(* IEC 61131-3 sources: iolistgen/pytests/golden/gen_fixture/src/POUs/Generated/PRG_Devices, 2 files *)

(* ---- PRG_Devices.decl.st ---- *)
// AUTO-GENERATED by iolistgen 0.2.0 — не редактировать; источник: gen_fixture.csv
// SHA-256 перечня 3ace79e7a28b; генератор st-codesys
// Назначение: вызовы устройств plc-process-lib по перечню сигналов: входы из GVL_IO, выходы в GVL_IO, команды GVL_Hmi,
// Cfg и Retain — GVL_Persist (контракт plc-process-lib, разделы 1 и 20). Входы автоматики (xAutoRun, xAutoOpen,
// wInterlock, wPermit…, rSpeedSpAuto_pct, rPosSpAuto_pct) пишет логика станции до вызова PRG_Devices; ПИД-регуляторы
// (тип Pid) без сигналов ввода-вывода вызывает логика станции (контракт 17.3)
// Автор:      iolistgen (генератор по перечню сигналов); перечень gen_fixture.csv
// Версия:     iolistgen 0.2.0
// Документ:   docs/signal_list.md
PROGRAM PRG_Devices
VAR
END_VAR

(* ---- PRG_Devices.impl.st ---- *)
// AUTO-GENERATED by iolistgen 0.2.0 — не редактировать; источник: gen_fixture.csv
// SHA-256 перечня 3ace79e7a28b; генератор st-codesys
// Порядок: устройства, на которые ссылаются link_power и link_fb (PWR2, ZT201), вызываются раньше ссылающихся; дальше —
// по dev_no.
// Источник времени не привязан: устройства берут встроенное системное время (контракт 20).

// Команда HMI «Применить уставки проекта» (контракт 18.3, правило 2): Retain устройств не меняется
IF GVL_Hmi.xApplyProjectCfg THEN
    GVL_Hmi.xApplyProjectCfg := FALSE;
    PRG_ApplyProjectCfg();
END_IF

// --- dev_no 6: PWR2 — Напряжение на секции шин (DigitalInput) ---
GVL_Devices.fbPWR2(
    xIn           := GVL_IO.xPWR2,
    xChannelFault := FALSE,  // нет строки CHF
    stCmd         := GVL_Hmi.stPWR2Cmd,
    stCfg         := GVL_Persist.stPWR2Cfg);

// --- dev_no 32: ZT201 — Клапан рециркуляции: положение (AnalogInput) ---
GVL_Devices.fbZT201(
    rIn           := GVL_IO.rZT201_mA,
    xChannelFault := FALSE,  // нет строки CHF
    stCmd         := GVL_Hmi.stZT201Cmd,
    stCfg         := GVL_Persist.stZT201Cfg);

// --- dev_no 1: LT201 — Уровень в резервуаре чистой воды (AnalogInput) ---
GVL_Devices.fbLT201(
    rIn           := GVL_IO.rLT201_mA,
    xChannelFault := GVL_IO.xLT201_CHF,
    stCmd         := GVL_Hmi.stLT201Cmd,
    stCfg         := GVL_Persist.stLT201Cfg);

// --- dev_no 2: PT201 — Давление на всасе (AnalogInput) ---
GVL_Devices.fbPT201(
    rIn           := INT_TO_REAL(GVL_IO.iPT201),
    xChannelFault := NOT GVL_IO.xMbOk_RS485_1_S5,  // нет строки CHF: обмен со слейвом
    stCmd         := GVL_Hmi.stPT201Cmd,
    stCfg         := GVL_Persist.stPT201Cfg);

// --- dev_no 3: TE201 — Температура воды (AnalogInput) ---
GVL_Devices.fbTE201(
    rIn           := GVL_IO.rTE201,
    xChannelFault := FALSE,  // нет строки CHF
    stCmd         := GVL_Hmi.stTE201Cmd,
    stCfg         := GVL_Persist.stTE201Cfg);

// --- dev_no 4: LS201 — Поплавок «перелив» (DigitalInput) ---
GVL_Devices.fbLS201(
    xIn           := GVL_IO.xLS201,
    xChannelFault := GVL_IO.xLS201_CHF,
    stCmd         := GVL_Hmi.stLS201Cmd,
    stCfg         := GVL_Persist.stLS201Cfg);

// --- dev_no 5: ES201 — Кнопка аварийного останова на щите (DigitalInput) ---
GVL_Devices.fbES201(
    xIn           := GVL_IO.xES201,
    xChannelFault := NOT GVL_IO.xMbOk_RS485_1_S7,  // нет строки CHF: обмен со слейвом
    stCmd         := GVL_Hmi.stES201Cmd,
    stCfg         := GVL_Persist.stES201Cfg);

// --- dev_no 11: M201 — Насос промывки (Motor) ---
GVL_Devices.fbM201(
    xFbRun    := GVL_IO.xM201_FB,
    xExtFault := GVL_IO.xM201_FLT,
    xLocal    := GVL_IO.xM201_LOC,
    xPowerOk  := GVL_Devices.fbPWR2.xValue,  // link_power
    stCmd     := GVL_Hmi.stM201Cmd,
    stCfg     := GVL_Persist.stM201Cfg,
    stRetain  := GVL_Persist.stM201Retain);
GVL_IO.xM201_RUN := GVL_Devices.fbM201.xQRun;
GVL_IO.xM201_RST := GVL_Devices.fbM201.xQReset;

// --- dev_no 12: P201 — Насос Н1 (MotorVfd) ---
// ПЧ: xCommOk, xVfd*, rSpeedAct_pct и rSpeedRef_pct — через адаптер приложения (GVL_IO.xP201_…)
GVL_Devices.fbP201(
    xExtFault     := GVL_IO.xP201_FLT,
    xLocal        := GVL_IO.xP201_LOC,
    xPowerOk      := GVL_Devices.fbPWR2.xValue,  // link_power
    xCommOk       := GVL_IO.xP201_CommOk,
    xVfdRunning   := GVL_IO.xP201_VfdRun,
    xVfdReady     := GVL_IO.xP201_VfdReady,
    xVfdFault     := GVL_IO.xP201_VfdFault,
    rSpeedAct_pct := GVL_IO.rP201_SpeedAct_pct,
    stCmd         := GVL_Hmi.stP201Cmd,
    stCfg         := GVL_Persist.stP201Cfg,
    stRetain      := GVL_Persist.stP201Retain);
GVL_IO.xP201_VfdQRun      := GVL_Devices.fbP201.xQRun;
GVL_IO.xP201_VfdQReset    := GVL_Devices.fbP201.xQReset;
GVL_IO.rP201_SpeedRef_pct := GVL_Devices.fbP201.rSpeedRef_pct;

// --- dev_no 13: P202 — Насос Н2 (MotorVfd) ---
// ПЧ: xCommOk, xVfd*, rSpeedAct_pct и rSpeedRef_pct — через адаптер приложения (GVL_IO.xP202_…)
GVL_Devices.fbP202(
    xFbRun        := GVL_IO.xP202_FB,
    xCommOk       := GVL_IO.xP202_CommOk,
    xVfdRunning   := GVL_IO.xP202_VfdRun,
    xVfdReady     := GVL_IO.xP202_VfdReady,
    xVfdFault     := GVL_IO.xP202_VfdFault,
    rSpeedAct_pct := GVL_IO.rP202_SpeedAct_pct,
    stCmd         := GVL_Hmi.stP202Cmd,
    stCfg         := GVL_Persist.stP202Cfg,
    stRetain      := GVL_Persist.stP202Retain);
GVL_IO.xP202_RUN          := GVL_Devices.fbP202.xQRun;
GVL_IO.rP202_SpeedRef_pct := GVL_Devices.fbP202.rSpeedRef_pct;

// --- dev_no 21: FV201 — Задвижка на напоре (Valve) ---
GVL_Devices.fbFV201(
    xZso         := GVL_IO.xFV201_ZSO,
    xZsc         := GVL_IO.xFV201_ZSC,
    xTorqueOpen  := GVL_IO.xFV201_TQO,
    xTorqueClose := GVL_IO.xFV201_TQC,
    xExtFault    := GVL_IO.xFV201_FLT,
    xLocal       := GVL_IO.xFV201_LOC,
    xPowerOk     := GVL_Devices.fbPWR2.xValue,  // link_power
    stCmd        := GVL_Hmi.stFV201Cmd,
    stCfg        := GVL_Persist.stFV201Cfg,
    stRetain     := GVL_Persist.stFV201Retain);
GVL_IO.xFV201_OPN := GVL_Devices.fbFV201.xQOpen;
GVL_IO.xFV201_CLS := GVL_Devices.fbFV201.xQClose;

// --- dev_no 22: XV201 — Клапан сброса (Valve) ---
GVL_Devices.fbXV201(
    xZsc     := GVL_IO.xXV201_ZSC,
    stCmd    := GVL_Hmi.stXV201Cmd,
    stCfg    := GVL_Persist.stXV201Cfg,
    stRetain := GVL_Persist.stXV201Retain);
GVL_IO.xXV201 := GVL_Devices.fbXV201.xQCoil;

// --- dev_no 31: FCV201 — Клапан рециркуляции (ControlValve) ---
GVL_Devices.fbFCV201(
    rPosFb_pct       := GVL_Devices.fbZT201.rValue_pct,  // link_fb
    xPosFbValid      := GVL_Devices.fbZT201.xValid,  // link_fb
    xLocal           := GVL_IO.xFCV201_LOC,
    xPositionerFault := GVL_IO.xFCV201_POSF,
    stCmd            := GVL_Hmi.stFCV201Cmd,
    stCfg            := GVL_Persist.stFCV201Cfg,
    stRetain         := GVL_Persist.stFCV201Retain);
GVL_IO.rFCV201_OUT_mA := GVL_Devices.fbFCV201.rOut_mA;

// --- dev_no 41: LIC201 — Регулятор уровня в резервуаре чистой воды (Pid) ---
// вызов FB_PID пишет логика станции до PRG_Devices (контракт plc-process-lib 17.3): входы rPv_eu, xPvValid, xTrack,
// rOutAct_pct и параметры ниже
// без входа ФБ (AUX, код приложения): GVL_IO.rLIC201_SPI — Регулятор уровня: задание на индикатор щита
// GVL_Devices.fbLIC201(
//     stCmd    := GVL_Hmi.stLIC201Cmd,
//     stCfg    := GVL_Persist.stLIC201Cfg,
//     stRetain := GVL_Persist.stLIC201Retain);
